Fanuc KAREL source: ks00047.KL

-- PROVISIONAL review KL for V1013-1; original PC SHA256 bb90b3ecf597ac1d93056bed6718a1cf430270f23cf3047ea0b22551668b5912
-- Incomplete behavior may be omitted. Consult companion uncertainty JSON. Do not deploy.
PROGRAM KS00047
%NOLOCKGROUP
BEGIN
  -- UNRESOLVED_PC offsets 5-13; opcodes 3F,75
  -- UNRESOLVED_PC offsets 18-27; opcodes 3F,75
  -- UNRESOLVED_PC offsets 32-45; opcodes 22,1D,23
  -- UNRESOLVED_PC offsets 50-54; opcodes 7F
END KS00047
